Fanuc KAREL source: ks00054.KL

PROGRAM KS00054
%STACKSIZE=65535
%PRIORITY=65535
%NOLOCKGROUP
TYPE
REC_T=STRUCTURE
VALUE : INTEGER
FLAG : BOOLEAN
ENDSTRUCTURE
VAR
A : ARRAY[4] OF REC_T
B : ARRAY[4] OF REC_T
FLAG : BOOLEAN
N : INTEGER
STATUS : INTEGER
PN : STRING[80]
VN : STRING[80]
BEGIN
PN=''
VN='A'
-- UNSAFE_SOURCE_IR line 19: N = native_s16_value(A)
END KS00054
